(* IEC 61131-3 sources: model-first-plc-agent-ai/pilot/reference, 4 files *)

(* ---- T1_ref.st ---- *)
(* Pilot reference program for task T1 (Factory I/O Scene 2, From A to B).
   For checking the compile script and the scene test before the formal run only:
   not a sample of RQ1 and not a listing of Section 5.2. *)

FUNCTION_BLOCK FB_FromAtoB
  VAR_INPUT
    sensor_a : BOOL;
    sensor_b : BOOL;
  END_VAR
  VAR_OUTPUT
    conveyor : BOOL;
  END_VAR
  VAR
    run_latch : RS;  (* reset dominant: a box at sensor B keeps the conveyor stopped *)
  END_VAR
  run_latch(S := sensor_a, R1 := sensor_b);
  conveyor := run_latch.Q1;
END_FUNCTION_BLOCK

PROGRAM Main
  VAR
    SensorA AT %IX100.0 : BOOL;
    SensorB AT %IX100.1 : BOOL;
    Conveyor AT %QX100.0 : BOOL;
  END_VAR
  VAR
    logic : FB_FromAtoB;
  END_VAR
  logic(sensor_a := SensorA, sensor_b := SensorB);
  Conveyor := logic.conveyor;
END_PROGRAM

(* ---- T2_ref.st ---- *)
(* Pilot reference program for task T2 (customized Scene 3, simple timer).
   For checking the compile script and the scene test before the formal run only:
   not a sample of RQ1 and not a listing of Section 5.2. *)

FUNCTION_BLOCK FB_SimpleTimerFill
  VAR_INPUT
    start_cmd : BOOL;
    stop_cmd : BOOL;
    lshh : BOOL;
    timer_duration : TIME;
  END_VAR
  VAR_OUTPUT
    fill_valve : BOOL;
    discharge_valve : BOOL;
  END_VAR
  VAR
    start_edge : R_TRIG;      (* start: TRUE only in the scan in which StartCommand is pressed *)
    fill_timer : TON;         (* timer of the filling step, IN := activity of step E1 *)
    x0 : BOOL := TRUE;        (* step 0 *)
    xe1 : BOOL := FALSE;      (* filling step E1 *)
  END_VAR
  start_edge(CLK := start_cmd);
  fill_timer(IN := xe1, PT := timer_duration);
  IF stop_cmd THEN
    x0 := TRUE;
    xe1 := FALSE;
  ELSIF x0 AND start_edge.Q THEN
    x0 := FALSE;
    xe1 := TRUE;
  ELSIF xe1 AND (fill_timer.Q OR lshh) THEN
    xe1 := FALSE;
    x0 := TRUE;
  END_IF;
  fill_valve := xe1;
  discharge_valve := FALSE;
END_FUNCTION_BLOCK

PROGRAM Main
  VAR
    StartCommand AT %IX100.0 : BOOL;
    StopCommand AT %IX100.1 : BOOL;
    LSH AT %IX100.2 : BOOL;
    LSHH AT %IX100.3 : BOOL;
    FillValve AT %QX100.0 : BOOL;
    DischargeValve AT %QX100.1 : BOOL;
  END_VAR
  VAR
    TimerDuration : TIME := T#15s;  (* scene test (a) T#15s: ends before LSH; (b) T#60s: LSHH ends filling *)
    logic : FB_SimpleTimerFill;
  END_VAR
  logic(start_cmd := StartCommand, stop_cmd := StopCommand, lshh := LSHH, timer_duration := TimerDuration);
  FillValve := logic.fill_valve;
  DischargeValve := logic.discharge_valve;
END_PROGRAM

(* ---- T3_ref.st ---- *)
(* Pilot reference program for task T3 (customized Scene 3, TON and TOF timers).
   For checking the compile script and the scene test before the formal run only:
   not a sample of RQ1 and not a listing of Section 5.2. *)

FUNCTION_BLOCK FB_TonTofFill
  VAR_INPUT
    start_cmd : BOOL;
    stop_cmd : BOOL;
    lsh : BOOL;
    ton_duration : TIME;
    tof_duration : TIME;
  END_VAR
  VAR_OUTPUT
    fill_valve : BOOL;
    discharge_valve : BOOL;
  END_VAR
  VAR
    start_edge : R_TRIG;
    ton_timer : TON;          (* IN := activity of filling step 21 *)
    tof_timer : TOF;          (* IN := activity of filling step 21; Q stays TRUE for tof_duration after step 21 is left *)
    x0 : BOOL := TRUE;        (* step 0 *)
    x21 : BOOL := FALSE;      (* filling step 21 *)
    x22 : BOOL := FALSE;      (* pause step 22 *)
  END_VAR
  start_edge(CLK := start_cmd);
  ton_timer(IN := x21, PT := ton_duration);
  tof_timer(IN := x21, PT := tof_duration);
  IF stop_cmd THEN
    x0 := TRUE;
    x21 := FALSE;
    x22 := FALSE;
  ELSIF x0 AND start_edge.Q THEN
    x0 := FALSE;
    x21 := TRUE;
  ELSIF x21 AND lsh THEN
    x21 := FALSE;
    x0 := TRUE;
  ELSIF x21 AND ton_timer.Q AND NOT lsh THEN
    x21 := FALSE;
    x22 := TRUE;
  ELSIF x22 AND NOT tof_timer.Q THEN
    x22 := FALSE;
    x21 := TRUE;
  END_IF;
  fill_valve := x21;
  discharge_valve := FALSE;
END_FUNCTION_BLOCK

PROGRAM Main
  VAR
    StartCommand AT %IX100.0 : BOOL;
    StopCommand AT %IX100.1 : BOOL;
    LSH AT %IX100.2 : BOOL;
    LSHH AT %IX100.3 : BOOL;
    FillValve AT %QX100.0 : BOOL;
    DischargeValve AT %QX100.1 : BOOL;
  END_VAR
  VAR
    TON_Duration : TIME := T#5s;
    TOF_Duration : TIME := T#5s;
    logic : FB_TonTofFill;
  END_VAR
  logic(start_cmd := StartCommand, stop_cmd := StopCommand, lsh := LSH,
        ton_duration := TON_Duration, tof_duration := TOF_Duration);
  FillValve := logic.fill_valve;
  DischargeValve := logic.discharge_valve;
END_PROGRAM

(* ---- T4_ref.st ---- *)
(* Pilot reference program for task T4 (Factory I/O Level Control, PID control).
   For checking the compile script and the scene test before the formal run only:
   not a sample of RQ1 and not a listing of Section 5.2.
   FULL_SCALE = 1000 as in the task card (Factory I/O Modbus TCP/IP Server driver with Scale = 100).
   Kp, Ti and Td come from pilot/pid_pretune.py and are confirmed by the logic analysis in pilot/vc
   (this program compiled and run in closed loop; frequency-domain margins).  They are not tuned in
   Factory I/O (author's ruling, 2026-11-13). *)

FUNCTION_BLOCK FB_LevelPID
  VAR_INPUT
    start_cmd : BOOL;
    stop_cmd : BOOL;
    level_raw : INT;
    full_scale : INT;
    kp : REAL;
    ti : REAL;          (* integral time in s; 0 disables the integral action *)
    td : REAL;          (* derivative time in s *)
    ts : REAL;          (* sampling period in s, equal to the task interval *)
  END_VAR
  VAR_OUTPUT
    fill_cmd : INT;
    discharge_cmd : INT;
  END_VAR
  VAR
    start_edge : R_TRIG;
    hold_timer : TON;   (* settled: |e| <= eps has held for t_h *)
    x0 : BOOL := TRUE;
    xe3 : BOOL := FALSE;
    h : REAL;           (* level as a fraction of the measuring span *)
    e : REAL;
    e_prev : REAL;
    i_term : REAL;
    d_term : REAL;
    u_raw : REAL;
    u : REAL;
    h_sp : REAL := 0.8;
    h_max : REAL := 0.9;
    eps : REAL := 0.02;
    t_h : TIME := T#10s;
    u_d : REAL := 0.4;  (* constant discharge-valve opening *)
  END_VAR
  start_edge(CLK := start_cmd);
  IF full_scale > 0 THEN
    h := INT_TO_REAL(level_raw) / INT_TO_REAL(full_scale);
  ELSE
    h := 0.0;
  END_IF;
  e := h_sp - h;
  hold_timer(IN := xe3 AND (ABS(e) <= eps), PT := t_h);
  IF stop_cmd THEN
    x0 := TRUE;
    xe3 := FALSE;
  ELSIF x0 AND start_edge.Q THEN
    x0 := FALSE;
    xe3 := TRUE;
    i_term := 0.0;
    e_prev := e;
  ELSIF xe3 AND (hold_timer.Q OR (h >= h_max)) THEN
    xe3 := FALSE;
    x0 := TRUE;
  END_IF;
  IF xe3 THEN
    d_term := 0.0;
    IF ts > 0.0 THEN
      d_term := kp * td * (e - e_prev) / ts;
    END_IF;
    u_raw := kp * e + i_term + d_term;
    IF u_raw > 1.0 THEN
      u := 1.0;                      (* clamped: integration suspended *)
    ELSIF u_raw < 0.0 THEN
      u := 0.0;                      (* clamped: integration suspended *)
    ELSE
      u := u_raw;
      IF ti > 0.0 THEN
        i_term := i_term + kp * ts / ti * e;
      END_IF;
    END_IF;
    e_prev := e;
    fill_cmd := REAL_TO_INT(u * INT_TO_REAL(full_scale));
    discharge_cmd := REAL_TO_INT(u_d * INT_TO_REAL(full_scale));
  ELSE
    u := 0.0;
    fill_cmd := 0;
    discharge_cmd := 0;
  END_IF;
END_FUNCTION_BLOCK

PROGRAM Main
  VAR
    StartCommand AT %IX100.0 : BOOL;
    StopCommand AT %IX100.1 : BOOL;
    LevelMeter AT %IW100 : INT;
    FillValve AT %QW100 : INT;
    DischargeValve AT %QW101 : INT;
  END_VAR
  VAR
    FULL_SCALE : INT := 1000;   (* register value at 10 V: driver Scale = 100, see the task card *)
    Kp : REAL := 5.0;           (* pid_pretune.py; confirmed by pilot/vc *)
    Ti : REAL := 40.0;
    Td : REAL := 0.0;
    Ts : REAL := 0.02;          (* equals the 20 ms task interval of the compile script *)
    ctrl : FB_LevelPID;
  END_VAR
  ctrl(start_cmd := StartCommand, stop_cmd := StopCommand, level_raw := LevelMeter,
       full_scale := FULL_SCALE, kp := Kp, ti := Ti, td := Td, ts := Ts);
  FillValve := ctrl.fill_cmd;
  DischargeValve := ctrl.discharge_cmd;
END_PROGRAM
